Fanuc KAREL source: kb00130.KL

PROGRAM KB00130
%STACKSIZE=65535
%PRIORITY=65535
%NOLOCKGROUP
VAR
P1 : INTEGER
P2 : INTEGER
P3 : BOOLEAN
BEGIN
P1=1
P2=1
P3=TRUE
PEND_SEMA(P1,P2,P3)
END KB00130
